// TIA Portal V20 export
// export: Created 2026-10-12T16:46:22.6823337Z, ExportSetting WithDefaults, DisplayName Totally Integrated Automation Portal, DisplayVersion V20 Update 6, DisplayName TIA Portal Openness, DisplayVersion V20 Update 6, DisplayName TIA Portal Version Control Interface, DisplayVersion V20 Update 6, DisplayName SINAMICS Startdrive Advanced, DisplayVersion V20 SP1 Update 2, DisplayName SINAMICS Startdrive G110M, G120, G120C, G120D, G120P, G115D, DisplayVersion V20 SP1 Update 2, DisplayName SINAMICS Startdrive G130, G150, S120, S150, SINAMICS MV, G220, S200, S210, DisplayVersion V20 SP1 Update 2, DisplayName STEP 7 Professional, DisplayVersion V20 Update 6, DisplayName STEP 7 Safety, DisplayVersion V20 Update 2, DisplayName WinCC Basic/Comfort/Advanced, DisplayVersion V20 Update 6, DisplayName WinCC Professional, DisplayVersion V20 Update 6, DisplayName WinCC Unified, DisplayVersion V20 Update 6
TYPE "UDT_KP8"
// stored: IsFailsafeCompliant false
   STRUCT
      Rohdaten : Struct
         IB_Tasten : Byte;
         IB_DI : Byte;
         QB_Rot : Byte;
         QB_Gruen : Byte;
         QB_Blau : Byte;
         QB_DO : Byte;
      END_STRUCT;
      Taste : Array[0..7] of Bool;
      LED : Array[0..7] of USInt;   // 0=Aus, 1=Rot, 2=Grün, 3=Blau, 4=Gelb, 5=Weiß
      DI : Array[0..7] of Bool;
      "DO" : Array[0..7] of Bool;
   END_STRUCT;
END_TYPE
